SYSTEM Filling2Module (* Module Filling2, generated from its module specification *)
  (* Standard: 61499-2 *)
  APPLICATION Filling2 (* Module Filling2 on target pc (localhost, IO modbus; generated by modgen) *)
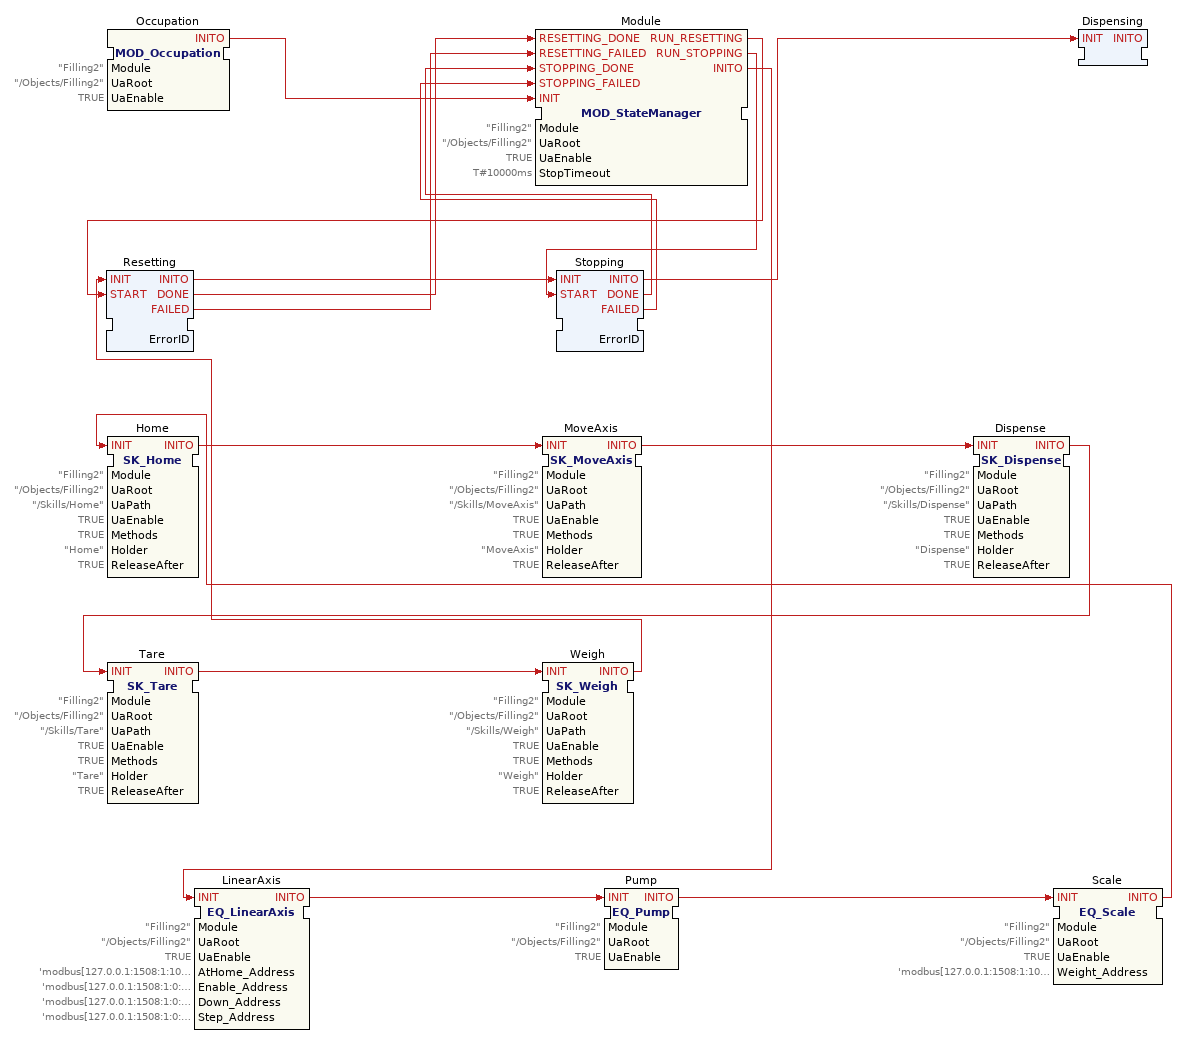
    (* Group ModuleLevel: Module level: occupation, PackML state manager, start-up and the target's IO lines *)
    (* Group ModuleLevelSkills: Module level skills: Control, Sequences (Execute, Stop) of skill primitives and Release; OPC UA /Skills/<name> *)
    (* Group Procedures: Procedures the module state manager runs while Resetting and Stopping *)
    (* Group SkillPrimitives: Skill primitives: one equipment command until a sensor or a time; OPC UA /Skills/<name> *)
    (* Group EquipmentIO: Equipment IO: the only owners of the IO points; skills send them output values over local channels *)
    FBS
      Occupation : modlib::MOD_Occupation(Module := "Filling2", UaRoot := "/Objects/Filling2", UaEnable := TRUE); (* Who may command the module. A client calls Occupy(Session) at /Objects/Filling2/Occupation first; until it calls Release, only commands with that session id are accepted. Every block hears the owner on loc[Filling2/owner]. *) {SET_ATTRIBUTE(GroupName, ModuleLevel)}
      Module : modlib::MOD_StateManager(Module := "Filling2", UaRoot := "/Objects/Filling2", UaEnable := TRUE, StopTimeout := T#10000ms); (* The module's PackML state. The owner calls Reset, Start, Stop, Abort or Clear at /Objects/Filling2/Module; State is at /Objects/Filling2/Module/State and on loc[Filling2/state]. Reset runs the Resetting procedure, Stop the Stopping procedure; skills may be started only in Execute. *) {SET_ATTRIBUTE(GroupName, ModuleLevel)}
      LinearAxis : filling::EQ_LinearAxis(Module := "Filling2", UaRoot := "/Objects/Filling2", UaEnable := TRUE, AtHome_Address := 'modbus[127.0.0.1:1508:1:10:d0:]', Enable_Address := 'modbus[127.0.0.1:1508:1:0::c0]', Down_Address := 'modbus[127.0.0.1:1508:1:0::c1]', Step_Address := 'modbus[127.0.0.1:1508:1:0::h0]'); (* Equipment LinearAxis: Needle lift, a stepper motor through a step and direction driver, with a limit switch at the top (home). The only block that touches its pins (AtHome = modbus[127.0.0.1:1508:1:10:d0:], Enable = modbus[127.0.0.1:1508:1:0::c0], Down = modbus[127.0.0.1:1508:1:0::c1], Step = modbus[127.0.0.1:1508:1:0::h0]). Skills send it what to switch on loc[Filling2/LinearAxis/cmd]; it reports its inputs on loc[Filling2/LinearAxis/state] and at /Objects/Filling2/Equipment/LinearAxis. *) {SET_ATTRIBUTE(GroupName, EquipmentIO)}
      Pump : filling::EQ_Pump(Module := "Filling2", UaRoot := "/Objects/Filling2", UaEnable := TRUE); (* Equipment Pump: Filling pump; none is wired yet, so it has no outputs and dispensing is a time at the station's flow rate. The only block that touches its pins (no pins). Skills send it what to switch on loc[Filling2/Pump/cmd]; it reports its inputs on loc[Filling2/Pump/state] and at /Objects/Filling2/Equipment/Pump. *) {SET_ATTRIBUTE(GroupName, EquipmentIO)}
      Scale : filling::EQ_Scale(Module := "Filling2", UaRoot := "/Objects/Filling2", UaEnable := TRUE, Weight_Address := 'modbus[127.0.0.1:1508:1:10:i0:]'); (* Equipment Scale: Scale; the hardware has none, so the weight is simulated. The only block that touches its pins (Weight = modbus[127.0.0.1:1508:1:10:i0:]). Skills send it what to switch on loc[Filling2/Scale/cmd]; it reports its inputs on loc[Filling2/Scale/state] and at /Objects/Filling2/Equipment/Scale. *) {SET_ATTRIBUTE(GroupName, EquipmentIO)}
      Home : filling::SK_Home(Module := "Filling2", UaRoot := "/Objects/Filling2", UaPath := "/Skills/Home", UaEnable := TRUE, Methods := TRUE, Holder := "Home", ReleaseAfter := TRUE); (* Skill Home, offered on its own: Needle up to the limit switch; from there its position is known, using LinearAxis. A client calls Start (with the parameters), Stop, Abort or Reset at /Objects/Filling2/Skills/Home; State, ErrorID, Parameters and Results are there too. *) {SET_ATTRIBUTE(GroupName, SkillPrimitives)}
      MoveAxis : filling::SK_MoveAxis(Module := "Filling2", UaRoot := "/Objects/Filling2", UaPath := "/Skills/MoveAxis", UaEnable := TRUE, Methods := TRUE, Holder := "MoveAxis", ReleaseAfter := TRUE); (* Skill MoveAxis, offered on its own: Needle to Position, measured down from the limit switch; the direction follows from where it is, using LinearAxis. A client calls Start (with the parameters), Stop, Abort or Reset at /Objects/Filling2/Skills/MoveAxis; State, ErrorID, Parameters and Results are there too. *) {SET_ATTRIBUTE(GroupName, SkillPrimitives)}
      Dispense : filling::SK_Dispense(Module := "Filling2", UaRoot := "/Objects/Filling2", UaPath := "/Skills/Dispense", UaEnable := TRUE, Methods := TRUE, Holder := "Dispense", ReleaseAfter := TRUE); (* Skill Dispense, offered on its own: Dispense a volume at the station's flow rate (open loop, by time, until a pump is wired), using Pump. A client calls Start (with the parameters), Stop, Abort or Reset at /Objects/Filling2/Skills/Dispense; State, ErrorID, Parameters and Results are there too. *) {SET_ATTRIBUTE(GroupName, SkillPrimitives)}
      Tare : filling::SK_Tare(Module := "Filling2", UaRoot := "/Objects/Filling2", UaPath := "/Skills/Tare", UaEnable := TRUE, Methods := TRUE, Holder := "Tare", ReleaseAfter := TRUE); (* Skill Tare, offered on its own: Tare the scale, using Scale. A client calls Start (with the parameters), Stop, Abort or Reset at /Objects/Filling2/Skills/Tare; State, ErrorID, Parameters and Results are there too. *) {SET_ATTRIBUTE(GroupName, SkillPrimitives)}
      Weigh : filling::SK_Weigh(Module := "Filling2", UaRoot := "/Objects/Filling2", UaPath := "/Skills/Weigh", UaEnable := TRUE, Methods := TRUE, Holder := "Weigh", ReleaseAfter := TRUE); (* Skill Weigh, offered on its own: Read the weight, using Scale. A client calls Start (with the parameters), Stop, Abort or Reset at /Objects/Filling2/Skills/Weigh; State, ErrorID, Parameters and Results are there too. *) {SET_ATTRIBUTE(GroupName, SkillPrimitives)}
    END_FBS
    SUBAPPLICATION Resetting (* Procedure the module runs while Resetting *)
      {SET_ATTRIBUTE(GroupName, Procedures)}
      EVENT_INPUT
        INIT : EInit;
        START;
      END_EVENT
      EVENT_OUTPUT
        INITO : EInit;
        DONE;
        FAILED;
      END_EVENT
      VAR_OUTPUT
        ErrorID : UINT;
      END_VAR
      FBS
        Home : filling::SK_Home(Module := "Filling2", UaRoot := "/Objects/Filling2", UaPath := "/Procedures/Resetting/Home", UaEnable := TRUE, Methods := FALSE, Holder := "Procedures/Resetting", ReleaseAfter := TRUE); (* Step 1 of Resetting: runs the skill Home. Its State and ErrorID are at /Objects/Filling2/Procedures/Resetting/Home; it keeps the equipment under the name Procedures/Resetting. *)
        Tare : filling::SK_Tare(Module := "Filling2", UaRoot := "/Objects/Filling2", UaPath := "/Procedures/Resetting/Tare", UaEnable := TRUE, Methods := FALSE, Holder := "Procedures/Resetting", ReleaseAfter := TRUE); (* Step 2 of Resetting: runs the skill Tare. Its State and ErrorID are at /Objects/Filling2/Procedures/Resetting/Tare; it keeps the equipment under the name Procedures/Resetting. *)
        Fail1 : modlib::SKILL_FailMerge; (* Joins the failures of the steps into one (with its error code), so any step's failure ends the sequence. *)
      END_FBS
      EVENT_CONNECTIONS
        Home.SUCCESS TO Tare.START;
        START TO Home.START;
        Tare.SUCCESS TO DONE;
        Home.FAILURE TO Fail1.FAIL_1;
        Tare.FAILURE TO Fail1.FAIL_2;
        Fail1.FAIL TO FAILED;
        INIT TO Home.INIT;
        Tare.INITO TO INITO;
        Home.INITO TO Tare.INIT;
      END_CONNECTIONS
      DATA_CONNECTIONS
        Home.ErrorID TO Fail1.Error1;
        Tare.ErrorID TO Fail1.Error2;
        Fail1.Error TO ErrorID;
      END_CONNECTIONS
    END_SUBAPPLICATION
    SUBAPPLICATION Stopping (* Procedure the module runs while Stopping *)
      {SET_ATTRIBUTE(GroupName, Procedures)}
      EVENT_INPUT
        INIT : EInit;
        START;
      END_EVENT
      EVENT_OUTPUT
        INITO : EInit;
        DONE;
        FAILED;
      END_EVENT
      VAR_OUTPUT
        ErrorID : UINT;
      END_VAR
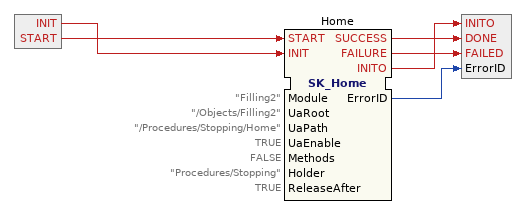
      FBS
        Home : filling::SK_Home(Module := "Filling2", UaRoot := "/Objects/Filling2", UaPath := "/Procedures/Stopping/Home", UaEnable := TRUE, Methods := FALSE, Holder := "Procedures/Stopping", ReleaseAfter := TRUE); (* Step 1 of Stopping: runs the skill Home. Its State and ErrorID are at /Objects/Filling2/Procedures/Stopping/Home; it keeps the equipment under the name Procedures/Stopping. *)
      END_FBS
      EVENT_CONNECTIONS
        START TO Home.START;
        Home.SUCCESS TO DONE;
        Home.FAILURE TO FAILED;
        INIT TO Home.INIT;
        Home.INITO TO INITO;
      END_CONNECTIONS
      DATA_CONNECTIONS
        Home.ErrorID TO ErrorID;
      END_CONNECTIONS
    END_SUBAPPLICATION
    SUBAPPLICATION Dispensing (* Module level skill Dispensing: Needle down, dispense the volume, needle up, weigh (runFillingCycle) *)
      {SET_ATTRIBUTE(GroupName, ModuleLevelSkills)}
      EVENT_INPUT
        INIT : EInit;
      END_EVENT
      EVENT_OUTPUT
        INITO : EInit;
      END_EVENT
      (* Group Core: The skill's state machine: Stop, Abort, Reset, State and ErrorID over OPC UA; gives up everything the skill holds when a run ends *)
      (* Group Start: The Start method: one block per parameter (range check, value for this run), the values published *)
      (* Group Sequences: What the skill does: Execute, and Stop when it is interrupted; private skill primitives in order *)
      (* Group Results: The results published when Execute is done *)
      FBS
        Control : modlib::SKILL_Core(Module := "Filling2", UaRoot := "/Objects/Filling2", UaPath := "/Skills/Dispensing", UaEnable := TRUE, Methods := TRUE, Holder := "Dispensing", ReleaseAll := TRUE); (* The state machine of the skill Dispensing: checks a client's Start (occupation, module in Execute, not running, values in range), publishes State and ErrorID at /Objects/Filling2/Skills/Dispensing, offers Stop, Abort and Reset there, starts Execute and runs Stop when the skill is stopped. *) {SET_ATTRIBUTE(GroupName, Core)}
        UaStart : iec61499::net::SERVER_2_2(QI := TRUE); (* The OPC UA method Start of Dispensing: a client's call (session id and parameters) arrives here; the parameters are checked, then Control answers Accepted or an error code. *) {SET_ATTRIBUTE(GroupName, Start)}
        Volume : modlib::SKILL_Param_LREAL(Default := 1.0, Lower := 0.5, Upper := 10.0); (* The parameter Volume of Dispensing: default 1.0 (Lower 0.5, Upper 10.0); checks a client's value, then holds it for the run and hands it to the steps. *) {SET_ATTRIBUTE(GroupName, Start)}
        PubParams : iec61499::net::PUBLISH_1(QI := TRUE, ID := "opc_ua[WRITE;/Objects/Filling2/Skills/Dispensing/Parameters/Volume]"); (* Writes the parameters of the run to OPC UA: /Objects/Filling2/Skills/Dispensing/Parameters/Volume *) {SET_ATTRIBUTE(GroupName, Start)}
        PubResults : iec61499::net::PUBLISH_1(QI := TRUE, ID := "opc_ua[WRITE;/Objects/Filling2/Skills/Dispensing/Results/Weight]"); (* Writes the results of the run to OPC UA: /Objects/Filling2/Skills/Dispensing/Results/Weight *) {SET_ATTRIBUTE(GroupName, Results)}
      END_FBS
      SUBAPPLICATION Execute (* Dispensing: execute sequence *)
        {SET_ATTRIBUTE(GroupName, Sequences)}
        EVENT_INPUT
          INIT : EInit;
          START;
          HALT;
          ABORT;
          RESET;
        END_EVENT
        EVENT_OUTPUT
          INITO : EInit;
          DONE;
          FAILED;
        END_EVENT
        VAR_INPUT
          Volume : LREAL;
        END_VAR
        VAR_OUTPUT
          ErrorID : UINT;
          Weight : LREAL;
        END_VAR
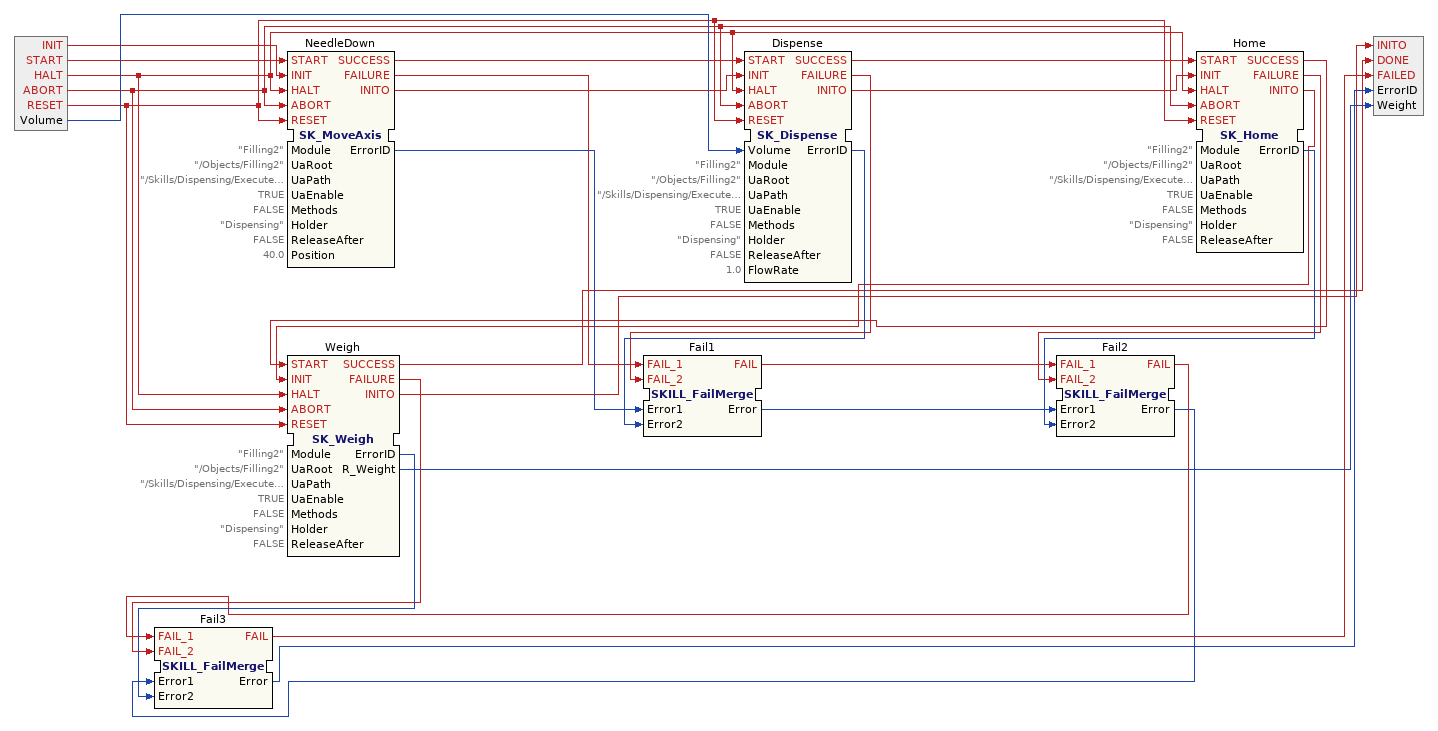
        FBS
          NeedleDown : filling::SK_MoveAxis(Module := "Filling2", UaRoot := "/Objects/Filling2", UaPath := "/Skills/Dispensing/Execute/NeedleDown", UaEnable := TRUE, Methods := FALSE, Holder := "Dispensing", ReleaseAfter := FALSE, Position := 40.0); (* Step 1 of Dispensing / Execute: runs the skill MoveAxis with Position = 40.0. Its State and ErrorID are at /Objects/Filling2/Skills/Dispensing/Execute/NeedleDown; it keeps the equipment under the name Dispensing. *)
          Dispense : filling::SK_Dispense(Module := "Filling2", UaRoot := "/Objects/Filling2", UaPath := "/Skills/Dispensing/Execute/Dispense", UaEnable := TRUE, Methods := FALSE, Holder := "Dispensing", ReleaseAfter := FALSE, FlowRate := 1.0); (* Step 2 of Dispensing / Execute: runs the skill Dispense with FlowRate = 1.0; Volume from Dispensing's Volume. Its State and ErrorID are at /Objects/Filling2/Skills/Dispensing/Execute/Dispense; it keeps the equipment under the name Dispensing. *)
          Home : filling::SK_Home(Module := "Filling2", UaRoot := "/Objects/Filling2", UaPath := "/Skills/Dispensing/Execute/Home", UaEnable := TRUE, Methods := FALSE, Holder := "Dispensing", ReleaseAfter := FALSE); (* Step 3 of Dispensing / Execute: runs the skill Home. Its State and ErrorID are at /Objects/Filling2/Skills/Dispensing/Execute/Home; it keeps the equipment under the name Dispensing. *)
          Weigh : filling::SK_Weigh(Module := "Filling2", UaRoot := "/Objects/Filling2", UaPath := "/Skills/Dispensing/Execute/Weigh", UaEnable := TRUE, Methods := FALSE, Holder := "Dispensing", ReleaseAfter := FALSE); (* Step 4 of Dispensing / Execute: runs the skill Weigh; its Weight is Dispensing's result. Its State and ErrorID are at /Objects/Filling2/Skills/Dispensing/Execute/Weigh; it keeps the equipment under the name Dispensing. *)
          Fail1 : modlib::SKILL_FailMerge; (* Joins the failures of the steps into one (with its error code), so any step's failure ends the sequence. *)
          Fail2 : modlib::SKILL_FailMerge; (* Joins the failures of the steps into one (with its error code), so any step's failure ends the sequence. *)
          Fail3 : modlib::SKILL_FailMerge; (* Joins the failures of the steps into one (with its error code), so any step's failure ends the sequence. *)
        END_FBS
        EVENT_CONNECTIONS
          NeedleDown.SUCCESS TO Dispense.START;
          Dispense.SUCCESS TO Home.START;
          Home.SUCCESS TO Weigh.START;
          START TO NeedleDown.START;
          Weigh.SUCCESS TO DONE;
          NeedleDown.FAILURE TO Fail1.FAIL_1;
          Dispense.FAILURE TO Fail1.FAIL_2;
          Fail1.FAIL TO Fail2.FAIL_1;
          Home.FAILURE TO Fail2.FAIL_2;
          Fail2.FAIL TO Fail3.FAIL_1;
          Weigh.FAILURE TO Fail3.FAIL_2;
          Fail3.FAIL TO FAILED;
          INIT TO NeedleDown.INIT;
          Weigh.INITO TO INITO;
          NeedleDown.INITO TO Dispense.INIT;
          Dispense.INITO TO Home.INIT;
          Home.INITO TO Weigh.INIT;
          HALT TO NeedleDown.HALT;
          HALT TO Dispense.HALT;
          HALT TO Home.HALT;
          HALT TO Weigh.HALT;
          ABORT TO NeedleDown.ABORT;
          ABORT TO Dispense.ABORT;
          ABORT TO Home.ABORT;
          ABORT TO Weigh.ABORT;
          RESET TO NeedleDown.RESET;
          RESET TO Dispense.RESET;
          RESET TO Home.RESET;
          RESET TO Weigh.RESET;
        END_CONNECTIONS
        DATA_CONNECTIONS
          Volume TO Dispense.Volume;
          NeedleDown.ErrorID TO Fail1.Error1;
          Dispense.ErrorID TO Fail1.Error2;
          Fail1.Error TO Fail2.Error1;
          Home.ErrorID TO Fail2.Error2;
          Fail2.Error TO Fail3.Error1;
          Weigh.ErrorID TO Fail3.Error2;
          Fail3.Error TO ErrorID;
          Weigh.R_Weight TO Weight;
        END_CONNECTIONS
      END_SUBAPPLICATION
      SUBAPPLICATION Stop (* Dispensing: stop sequence *)
        {SET_ATTRIBUTE(GroupName, Sequences)}
        EVENT_INPUT
          INIT : EInit;
          START;
          HALT;
          ABORT;
          RESET;
        END_EVENT
        EVENT_OUTPUT
          INITO : EInit;
          DONE;
          FAILED;
        END_EVENT
        VAR_OUTPUT
          ErrorID : UINT;
        END_VAR
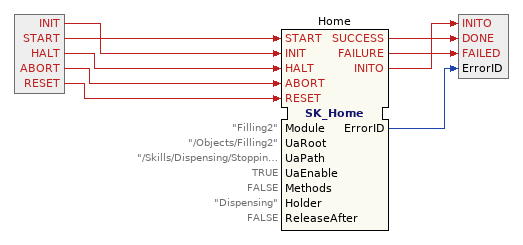
        FBS
          Home : filling::SK_Home(Module := "Filling2", UaRoot := "/Objects/Filling2", UaPath := "/Skills/Dispensing/Stopping/Home", UaEnable := TRUE, Methods := FALSE, Holder := "Dispensing", ReleaseAfter := FALSE); (* Step 1 of Dispensing / Stop: runs the skill Home. Its State and ErrorID are at /Objects/Filling2/Skills/Dispensing/Stopping/Home; it keeps the equipment under the name Dispensing. *)
        END_FBS
        EVENT_CONNECTIONS
          START TO Home.START;
          Home.SUCCESS TO DONE;
          Home.FAILURE TO FAILED;
          INIT TO Home.INIT;
          Home.INITO TO INITO;
          HALT TO Home.HALT;
          ABORT TO Home.ABORT;
          RESET TO Home.RESET;
        END_CONNECTIONS
        DATA_CONNECTIONS
          Home.ErrorID TO ErrorID;
        END_CONNECTIONS
      END_SUBAPPLICATION
      EVENT_CONNECTIONS
        Control.START_RSP TO UaStart.RSP;
        UaStart.IND TO Volume.CHECK;
        Control.RUN TO Volume.LATCH;
        Volume.CHECKED TO Control.START_REQ;
        Volume.LATCHED TO PubParams.REQ;
        PubParams.INITO TO PubParams.REQ;
        Execute.DONE TO PubResults.REQ;
        Volume.LATCHED TO Execute.START;
        Control.HALT_SEQ TO Execute.HALT;
        Control.ABORT_SEQ TO Execute.ABORT;
        Control.RESET_SEQ TO Execute.RESET;
        Execute.DONE TO Control.EXECUTE_DONE;
        Execute.FAILED TO Control.EXECUTE_FAILED;
        Control.RUN_STOPPING TO Stop.START;
        Control.ABORT_SEQ TO Stop.ABORT;
        Control.RESET_SEQ TO Stop.RESET;
        Stop.DONE TO Control.STOPPING_DONE;
        Stop.FAILED TO Control.STOPPING_DONE;
        INIT TO Control.INIT;
        Control.INITO TO UaStart.INIT;
        UaStart.INITO TO Volume.INIT;
        Volume.INITO TO PubParams.INIT;
        PubParams.INITO TO PubResults.INIT;
        PubResults.INITO TO Execute.INIT;
        Execute.INITO TO Stop.INIT;
        Stop.INITO TO INITO;
      END_CONNECTIONS
      DATA_CONNECTIONS
        Control.StartMethodId TO UaStart.ID;
        UaStart.RD_1 TO Control.Session;
        Control.Accepted TO UaStart.SD_1;
        Control.StartError TO UaStart.SD_2;
        UaStart.RD_2 TO Volume.Requested;
        Control.CalledByClient TO Volume.CalledByClient;
        Volume.Value TO PubParams.SD_1;
        Volume.AllInRange TO Control.ParamsInRange;
        Execute.Weight TO PubResults.SD_1;
        Volume.Value TO Execute.Volume;
        Execute.ErrorID TO Control.ExecuteError;
      END_CONNECTIONS
    END_SUBAPPLICATION
    EVENT_CONNECTIONS
      Module.RUN_RESETTING TO Resetting.START;
      Resetting.DONE TO Module.RESETTING_DONE;
      Resetting.FAILED TO Module.RESETTING_FAILED;
      Module.RUN_STOPPING TO Stopping.START;
      Stopping.DONE TO Module.STOPPING_DONE;
      Stopping.FAILED TO Module.STOPPING_FAILED;
      Occupation.INITO TO Module.INIT;
      Module.INITO TO LinearAxis.INIT;
      LinearAxis.INITO TO Pump.INIT;
      Pump.INITO TO Scale.INIT;
      Scale.INITO TO Home.INIT;
      Home.INITO TO MoveAxis.INIT;
      MoveAxis.INITO TO Dispense.INIT;
      Dispense.INITO TO Tare.INIT;
      Tare.INITO TO Weigh.INIT;
      Weigh.INITO TO Resetting.INIT;
      Resetting.INITO TO Stopping.INIT;
      Stopping.INITO TO Dispensing.INIT;
    END_CONNECTIONS
  END_APPLICATION
  APPLICATION Filling2_pi (* Module Filling2 on target pi (192.168.0.173, IO gpio; generated by modgen) *)
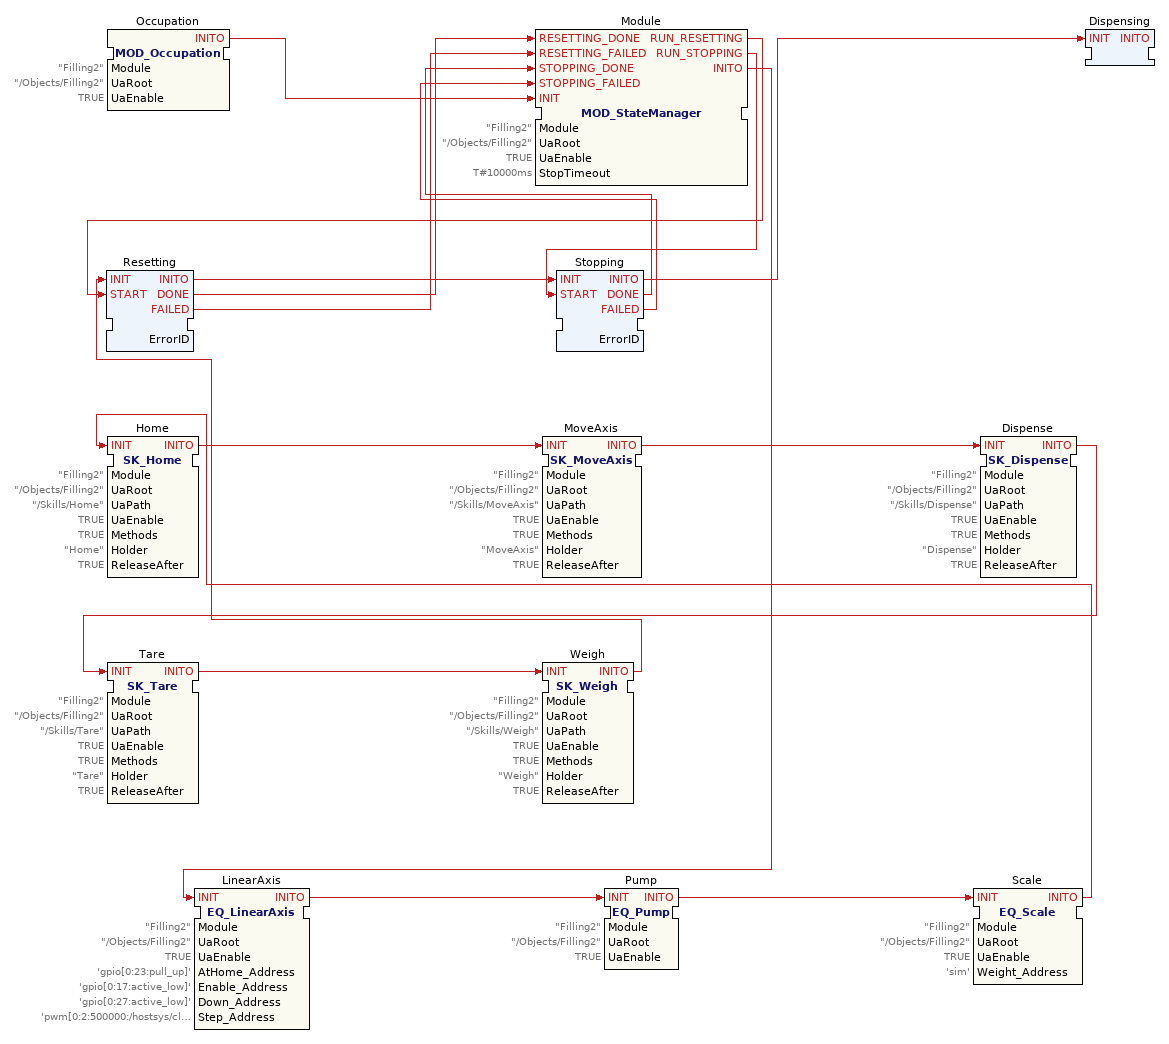
    (* Group ModuleLevel: Module level: occupation, PackML state manager, start-up and the target's IO lines *)
    (* Group ModuleLevelSkills: Module level skills: Control, Sequences (Execute, Stop) of skill primitives and Release; OPC UA /Skills/<name> *)
    (* Group Procedures: Procedures the module state manager runs while Resetting and Stopping *)
    (* Group SkillPrimitives: Skill primitives: one equipment command until a sensor or a time; OPC UA /Skills/<name> *)
    (* Group EquipmentIO: Equipment IO: the only owners of the IO points; skills send them output values over local channels *)
    FBS
      Occupation : modlib::MOD_Occupation(Module := "Filling2", UaRoot := "/Objects/Filling2", UaEnable := TRUE); (* Who may command the module. A client calls Occupy(Session) at /Objects/Filling2/Occupation first; until it calls Release, only commands with that session id are accepted. Every block hears the owner on loc[Filling2/owner]. *) {SET_ATTRIBUTE(GroupName, ModuleLevel)}
      Module : modlib::MOD_StateManager(Module := "Filling2", UaRoot := "/Objects/Filling2", UaEnable := TRUE, StopTimeout := T#10000ms); (* The module's PackML state. The owner calls Reset, Start, Stop, Abort or Clear at /Objects/Filling2/Module; State is at /Objects/Filling2/Module/State and on loc[Filling2/state]. Reset runs the Resetting procedure, Stop the Stopping procedure; skills may be started only in Execute. *) {SET_ATTRIBUTE(GroupName, ModuleLevel)}
      LinearAxis : filling::EQ_LinearAxis(Module := "Filling2", UaRoot := "/Objects/Filling2", UaEnable := TRUE, AtHome_Address := 'gpio[0:23:pull_up]', Enable_Address := 'gpio[0:17:active_low]', Down_Address := 'gpio[0:27:active_low]', Step_Address := 'pwm[0:2:500000:/hostsys/class/pwm]'); (* Equipment LinearAxis: Needle lift, a stepper motor through a step and direction driver, with a limit switch at the top (home). The only block that touches its pins (AtHome = gpio[0:23:pull_up], Enable = gpio[0:17:active_low], Down = gpio[0:27:active_low], Step = pwm[0:2:500000:/hostsys/class/pwm]). Skills send it what to switch on loc[Filling2/LinearAxis/cmd]; it reports its inputs on loc[Filling2/LinearAxis/state] and at /Objects/Filling2/Equipment/LinearAxis. *) {SET_ATTRIBUTE(GroupName, EquipmentIO)}
      Pump : filling::EQ_Pump(Module := "Filling2", UaRoot := "/Objects/Filling2", UaEnable := TRUE); (* Equipment Pump: Filling pump; none is wired yet, so it has no outputs and dispensing is a time at the station's flow rate. The only block that touches its pins (no pins). Skills send it what to switch on loc[Filling2/Pump/cmd]; it reports its inputs on loc[Filling2/Pump/state] and at /Objects/Filling2/Equipment/Pump. *) {SET_ATTRIBUTE(GroupName, EquipmentIO)}
      Scale : filling::EQ_Scale(Module := "Filling2", UaRoot := "/Objects/Filling2", UaEnable := TRUE, Weight_Address := 'sim'); (* Equipment Scale: Scale; the hardware has none, so the weight is simulated. The only block that touches its pins (Weight = sim). Skills send it what to switch on loc[Filling2/Scale/cmd]; it reports its inputs on loc[Filling2/Scale/state] and at /Objects/Filling2/Equipment/Scale. *) {SET_ATTRIBUTE(GroupName, EquipmentIO)}
      Home : filling::SK_Home(Module := "Filling2", UaRoot := "/Objects/Filling2", UaPath := "/Skills/Home", UaEnable := TRUE, Methods := TRUE, Holder := "Home", ReleaseAfter := TRUE); (* Skill Home, offered on its own: Needle up to the limit switch; from there its position is known, using LinearAxis. A client calls Start (with the parameters), Stop, Abort or Reset at /Objects/Filling2/Skills/Home; State, ErrorID, Parameters and Results are there too. *) {SET_ATTRIBUTE(GroupName, SkillPrimitives)}
      MoveAxis : filling::SK_MoveAxis(Module := "Filling2", UaRoot := "/Objects/Filling2", UaPath := "/Skills/MoveAxis", UaEnable := TRUE, Methods := TRUE, Holder := "MoveAxis", ReleaseAfter := TRUE); (* Skill MoveAxis, offered on its own: Needle to Position, measured down from the limit switch; the direction follows from where it is, using LinearAxis. A client calls Start (with the parameters), Stop, Abort or Reset at /Objects/Filling2/Skills/MoveAxis; State, ErrorID, Parameters and Results are there too. *) {SET_ATTRIBUTE(GroupName, SkillPrimitives)}
      Dispense : filling::SK_Dispense(Module := "Filling2", UaRoot := "/Objects/Filling2", UaPath := "/Skills/Dispense", UaEnable := TRUE, Methods := TRUE, Holder := "Dispense", ReleaseAfter := TRUE); (* Skill Dispense, offered on its own: Dispense a volume at the station's flow rate (open loop, by time, until a pump is wired), using Pump. A client calls Start (with the parameters), Stop, Abort or Reset at /Objects/Filling2/Skills/Dispense; State, ErrorID, Parameters and Results are there too. *) {SET_ATTRIBUTE(GroupName, SkillPrimitives)}
      Tare : filling::SK_Tare(Module := "Filling2", UaRoot := "/Objects/Filling2", UaPath := "/Skills/Tare", UaEnable := TRUE, Methods := TRUE, Holder := "Tare", ReleaseAfter := TRUE); (* Skill Tare, offered on its own: Tare the scale, using Scale. A client calls Start (with the parameters), Stop, Abort or Reset at /Objects/Filling2/Skills/Tare; State, ErrorID, Parameters and Results are there too. *) {SET_ATTRIBUTE(GroupName, SkillPrimitives)}
      Weigh : filling::SK_Weigh(Module := "Filling2", UaRoot := "/Objects/Filling2", UaPath := "/Skills/Weigh", UaEnable := TRUE, Methods := TRUE, Holder := "Weigh", ReleaseAfter := TRUE); (* Skill Weigh, offered on its own: Read the weight, using Scale. A client calls Start (with the parameters), Stop, Abort or Reset at /Objects/Filling2/Skills/Weigh; State, ErrorID, Parameters and Results are there too. *) {SET_ATTRIBUTE(GroupName, SkillPrimitives)}
    END_FBS
    SUBAPPLICATION Resetting (* Procedure the module runs while Resetting *)
      {SET_ATTRIBUTE(GroupName, Procedures)}
      EVENT_INPUT
        INIT : EInit;
        START;
      END_EVENT
      EVENT_OUTPUT
        INITO : EInit;
        DONE;
        FAILED;
      END_EVENT
      VAR_OUTPUT
        ErrorID : UINT;
      END_VAR
      FBS
        Home : filling::SK_Home(Module := "Filling2", UaRoot := "/Objects/Filling2", UaPath := "/Procedures/Resetting/Home", UaEnable := TRUE, Methods := FALSE, Holder := "Procedures/Resetting", ReleaseAfter := TRUE); (* Step 1 of Resetting: runs the skill Home. Its State and ErrorID are at /Objects/Filling2/Procedures/Resetting/Home; it keeps the equipment under the name Procedures/Resetting. *)
        Tare : filling::SK_Tare(Module := "Filling2", UaRoot := "/Objects/Filling2", UaPath := "/Procedures/Resetting/Tare", UaEnable := TRUE, Methods := FALSE, Holder := "Procedures/Resetting", ReleaseAfter := TRUE); (* Step 2 of Resetting: runs the skill Tare. Its State and ErrorID are at /Objects/Filling2/Procedures/Resetting/Tare; it keeps the equipment under the name Procedures/Resetting. *)
        Fail1 : modlib::SKILL_FailMerge; (* Joins the failures of the steps into one (with its error code), so any step's failure ends the sequence. *)
      END_FBS
      EVENT_CONNECTIONS
        Home.SUCCESS TO Tare.START;
        START TO Home.START;
        Tare.SUCCESS TO DONE;
        Home.FAILURE TO Fail1.FAIL_1;
        Tare.FAILURE TO Fail1.FAIL_2;
        Fail1.FAIL TO FAILED;
        INIT TO Home.INIT;
        Tare.INITO TO INITO;
        Home.INITO TO Tare.INIT;
      END_CONNECTIONS
      DATA_CONNECTIONS
        Home.ErrorID TO Fail1.Error1;
        Tare.ErrorID TO Fail1.Error2;
        Fail1.Error TO ErrorID;
      END_CONNECTIONS
    END_SUBAPPLICATION
    SUBAPPLICATION Stopping (* Procedure the module runs while Stopping *)
      {SET_ATTRIBUTE(GroupName, Procedures)}
      EVENT_INPUT
        INIT : EInit;
        START;
      END_EVENT
      EVENT_OUTPUT
        INITO : EInit;
        DONE;
        FAILED;
      END_EVENT
      VAR_OUTPUT
        ErrorID : UINT;
      END_VAR
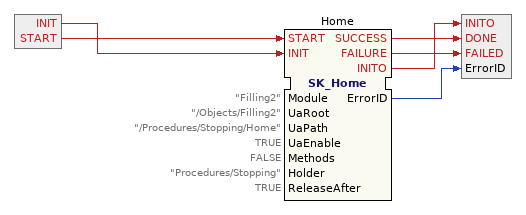
      FBS
        Home : filling::SK_Home(Module := "Filling2", UaRoot := "/Objects/Filling2", UaPath := "/Procedures/Stopping/Home", UaEnable := TRUE, Methods := FALSE, Holder := "Procedures/Stopping", ReleaseAfter := TRUE); (* Step 1 of Stopping: runs the skill Home. Its State and ErrorID are at /Objects/Filling2/Procedures/Stopping/Home; it keeps the equipment under the name Procedures/Stopping. *)
      END_FBS
      EVENT_CONNECTIONS
        START TO Home.START;
        Home.SUCCESS TO DONE;
        Home.FAILURE TO FAILED;
        INIT TO Home.INIT;
        Home.INITO TO INITO;
      END_CONNECTIONS
      DATA_CONNECTIONS
        Home.ErrorID TO ErrorID;
      END_CONNECTIONS
    END_SUBAPPLICATION
    SUBAPPLICATION Dispensing (* Module level skill Dispensing: Needle down, dispense the volume, needle up, weigh (runFillingCycle) *)
      {SET_ATTRIBUTE(GroupName, ModuleLevelSkills)}
      EVENT_INPUT
        INIT : EInit;
      END_EVENT
      EVENT_OUTPUT
        INITO : EInit;
      END_EVENT
      (* Group Core: The skill's state machine: Stop, Abort, Reset, State and ErrorID over OPC UA; gives up everything the skill holds when a run ends *)
      (* Group Start: The Start method: one block per parameter (range check, value for this run), the values published *)
      (* Group Sequences: What the skill does: Execute, and Stop when it is interrupted; private skill primitives in order *)
      (* Group Results: The results published when Execute is done *)
      FBS
        Control : modlib::SKILL_Core(Module := "Filling2", UaRoot := "/Objects/Filling2", UaPath := "/Skills/Dispensing", UaEnable := TRUE, Methods := TRUE, Holder := "Dispensing", ReleaseAll := TRUE); (* The state machine of the skill Dispensing: checks a client's Start (occupation, module in Execute, not running, values in range), publishes State and ErrorID at /Objects/Filling2/Skills/Dispensing, offers Stop, Abort and Reset there, starts Execute and runs Stop when the skill is stopped. *) {SET_ATTRIBUTE(GroupName, Core)}
        UaStart : iec61499::net::SERVER_2_2(QI := TRUE); (* The OPC UA method Start of Dispensing: a client's call (session id and parameters) arrives here; the parameters are checked, then Control answers Accepted or an error code. *) {SET_ATTRIBUTE(GroupName, Start)}
        Volume : modlib::SKILL_Param_LREAL(Default := 1.0, Lower := 0.5, Upper := 10.0); (* The parameter Volume of Dispensing: default 1.0 (Lower 0.5, Upper 10.0); checks a client's value, then holds it for the run and hands it to the steps. *) {SET_ATTRIBUTE(GroupName, Start)}
        PubParams : iec61499::net::PUBLISH_1(QI := TRUE, ID := "opc_ua[WRITE;/Objects/Filling2/Skills/Dispensing/Parameters/Volume]"); (* Writes the parameters of the run to OPC UA: /Objects/Filling2/Skills/Dispensing/Parameters/Volume *) {SET_ATTRIBUTE(GroupName, Start)}
        PubResults : iec61499::net::PUBLISH_1(QI := TRUE, ID := "opc_ua[WRITE;/Objects/Filling2/Skills/Dispensing/Results/Weight]"); (* Writes the results of the run to OPC UA: /Objects/Filling2/Skills/Dispensing/Results/Weight *) {SET_ATTRIBUTE(GroupName, Results)}
      END_FBS
      SUBAPPLICATION Execute (* Dispensing: execute sequence *)
        {SET_ATTRIBUTE(GroupName, Sequences)}
        EVENT_INPUT
          INIT : EInit;
          START;
          HALT;
          ABORT;
          RESET;
        END_EVENT
        EVENT_OUTPUT
          INITO : EInit;
          DONE;
          FAILED;
        END_EVENT
        VAR_INPUT
          Volume : LREAL;
        END_VAR
        VAR_OUTPUT
          ErrorID : UINT;
          Weight : LREAL;
        END_VAR
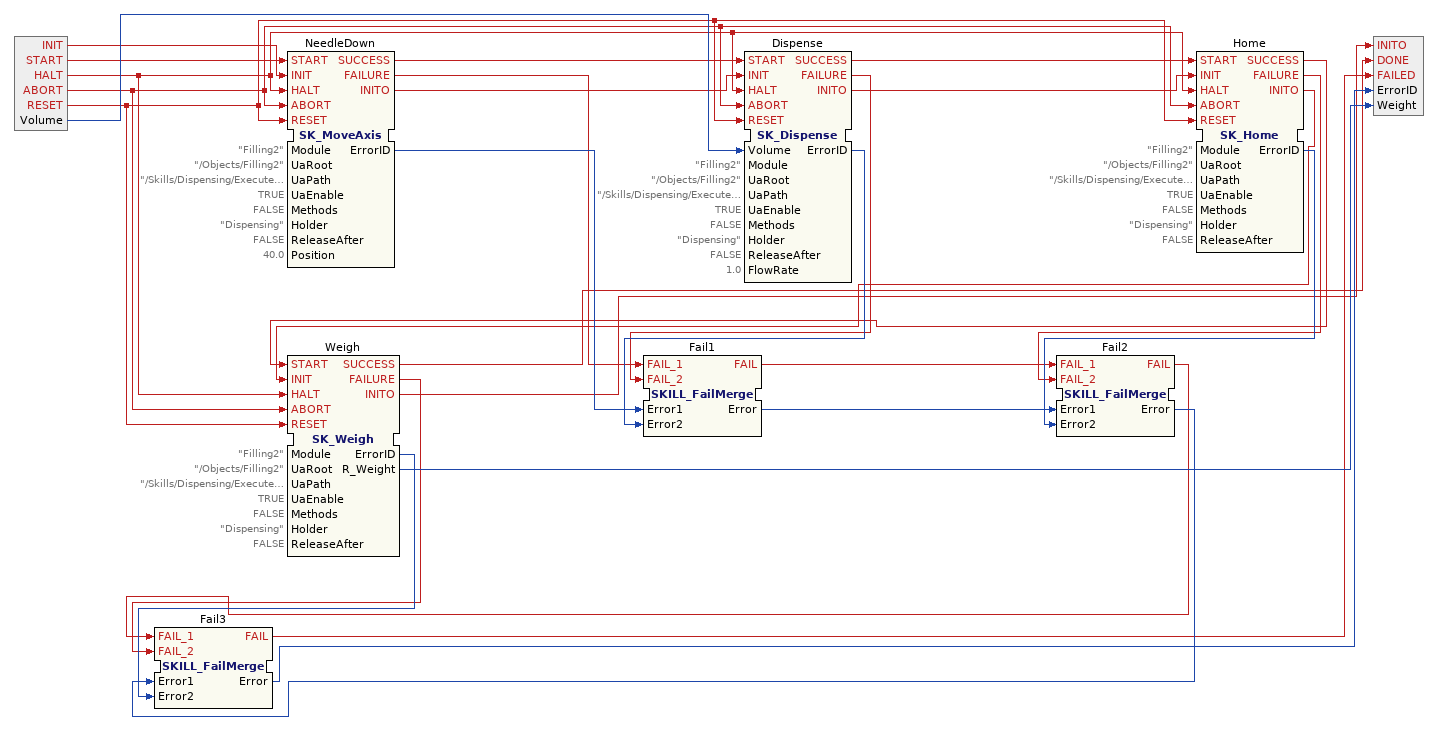
        FBS
          NeedleDown : filling::SK_MoveAxis(Module := "Filling2", UaRoot := "/Objects/Filling2", UaPath := "/Skills/Dispensing/Execute/NeedleDown", UaEnable := TRUE, Methods := FALSE, Holder := "Dispensing", ReleaseAfter := FALSE, Position := 40.0); (* Step 1 of Dispensing / Execute: runs the skill MoveAxis with Position = 40.0. Its State and ErrorID are at /Objects/Filling2/Skills/Dispensing/Execute/NeedleDown; it keeps the equipment under the name Dispensing. *)
          Dispense : filling::SK_Dispense(Module := "Filling2", UaRoot := "/Objects/Filling2", UaPath := "/Skills/Dispensing/Execute/Dispense", UaEnable := TRUE, Methods := FALSE, Holder := "Dispensing", ReleaseAfter := FALSE, FlowRate := 1.0); (* Step 2 of Dispensing / Execute: runs the skill Dispense with FlowRate = 1.0; Volume from Dispensing's Volume. Its State and ErrorID are at /Objects/Filling2/Skills/Dispensing/Execute/Dispense; it keeps the equipment under the name Dispensing. *)
          Home : filling::SK_Home(Module := "Filling2", UaRoot := "/Objects/Filling2", UaPath := "/Skills/Dispensing/Execute/Home", UaEnable := TRUE, Methods := FALSE, Holder := "Dispensing", ReleaseAfter := FALSE); (* Step 3 of Dispensing / Execute: runs the skill Home. Its State and ErrorID are at /Objects/Filling2/Skills/Dispensing/Execute/Home; it keeps the equipment under the name Dispensing. *)
          Weigh : filling::SK_Weigh(Module := "Filling2", UaRoot := "/Objects/Filling2", UaPath := "/Skills/Dispensing/Execute/Weigh", UaEnable := TRUE, Methods := FALSE, Holder := "Dispensing", ReleaseAfter := FALSE); (* Step 4 of Dispensing / Execute: runs the skill Weigh; its Weight is Dispensing's result. Its State and ErrorID are at /Objects/Filling2/Skills/Dispensing/Execute/Weigh; it keeps the equipment under the name Dispensing. *)
          Fail1 : modlib::SKILL_FailMerge; (* Joins the failures of the steps into one (with its error code), so any step's failure ends the sequence. *)
          Fail2 : modlib::SKILL_FailMerge; (* Joins the failures of the steps into one (with its error code), so any step's failure ends the sequence. *)
          Fail3 : modlib::SKILL_FailMerge; (* Joins the failures of the steps into one (with its error code), so any step's failure ends the sequence. *)
        END_FBS
        EVENT_CONNECTIONS
          NeedleDown.SUCCESS TO Dispense.START;
          Dispense.SUCCESS TO Home.START;
          Home.SUCCESS TO Weigh.START;
          START TO NeedleDown.START;
          Weigh.SUCCESS TO DONE;
          NeedleDown.FAILURE TO Fail1.FAIL_1;
          Dispense.FAILURE TO Fail1.FAIL_2;
          Fail1.FAIL TO Fail2.FAIL_1;
          Home.FAILURE TO Fail2.FAIL_2;
          Fail2.FAIL TO Fail3.FAIL_1;
          Weigh.FAILURE TO Fail3.FAIL_2;
          Fail3.FAIL TO FAILED;
          INIT TO NeedleDown.INIT;
          Weigh.INITO TO INITO;
          NeedleDown.INITO TO Dispense.INIT;
          Dispense.INITO TO Home.INIT;
          Home.INITO TO Weigh.INIT;
          HALT TO NeedleDown.HALT;
          HALT TO Dispense.HALT;
          HALT TO Home.HALT;
          HALT TO Weigh.HALT;
          ABORT TO NeedleDown.ABORT;
          ABORT TO Dispense.ABORT;
          ABORT TO Home.ABORT;
          ABORT TO Weigh.ABORT;
          RESET TO NeedleDown.RESET;
          RESET TO Dispense.RESET;
          RESET TO Home.RESET;
          RESET TO Weigh.RESET;
        END_CONNECTIONS
        DATA_CONNECTIONS
          Volume TO Dispense.Volume;
          NeedleDown.ErrorID TO Fail1.Error1;
          Dispense.ErrorID TO Fail1.Error2;
          Fail1.Error TO Fail2.Error1;
          Home.ErrorID TO Fail2.Error2;
          Fail2.Error TO Fail3.Error1;
          Weigh.ErrorID TO Fail3.Error2;
          Fail3.Error TO ErrorID;
          Weigh.R_Weight TO Weight;
        END_CONNECTIONS
      END_SUBAPPLICATION
      SUBAPPLICATION Stop (* Dispensing: stop sequence *)
        {SET_ATTRIBUTE(GroupName, Sequences)}
        EVENT_INPUT
          INIT : EInit;
          START;
          HALT;
          ABORT;
          RESET;
        END_EVENT
        EVENT_OUTPUT
          INITO : EInit;
          DONE;
          FAILED;
        END_EVENT
        VAR_OUTPUT
          ErrorID : UINT;
        END_VAR
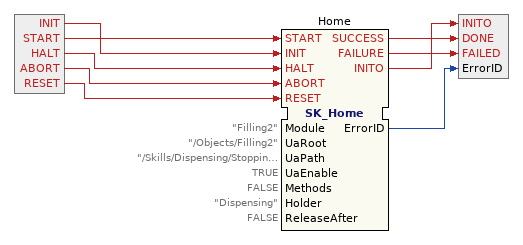
        FBS
          Home : filling::SK_Home(Module := "Filling2", UaRoot := "/Objects/Filling2", UaPath := "/Skills/Dispensing/Stopping/Home", UaEnable := TRUE, Methods := FALSE, Holder := "Dispensing", ReleaseAfter := FALSE); (* Step 1 of Dispensing / Stop: runs the skill Home. Its State and ErrorID are at /Objects/Filling2/Skills/Dispensing/Stopping/Home; it keeps the equipment under the name Dispensing. *)
        END_FBS
        EVENT_CONNECTIONS
          START TO Home.START;
          Home.SUCCESS TO DONE;
          Home.FAILURE TO FAILED;
          INIT TO Home.INIT;
          Home.INITO TO INITO;
          HALT TO Home.HALT;
          ABORT TO Home.ABORT;
          RESET TO Home.RESET;
        END_CONNECTIONS
        DATA_CONNECTIONS
          Home.ErrorID TO ErrorID;
        END_CONNECTIONS
      END_SUBAPPLICATION
      EVENT_CONNECTIONS
        Control.START_RSP TO UaStart.RSP;
        UaStart.IND TO Volume.CHECK;
        Control.RUN TO Volume.LATCH;
        Volume.CHECKED TO Control.START_REQ;
        Volume.LATCHED TO PubParams.REQ;
        PubParams.INITO TO PubParams.REQ;
        Execute.DONE TO PubResults.REQ;
        Volume.LATCHED TO Execute.START;
        Control.HALT_SEQ TO Execute.HALT;
        Control.ABORT_SEQ TO Execute.ABORT;
        Control.RESET_SEQ TO Execute.RESET;
        Execute.DONE TO Control.EXECUTE_DONE;
        Execute.FAILED TO Control.EXECUTE_FAILED;
        Control.RUN_STOPPING TO Stop.START;
        Control.ABORT_SEQ TO Stop.ABORT;
        Control.RESET_SEQ TO Stop.RESET;
        Stop.DONE TO Control.STOPPING_DONE;
        Stop.FAILED TO Control.STOPPING_DONE;
        INIT TO Control.INIT;
        Control.INITO TO UaStart.INIT;
        UaStart.INITO TO Volume.INIT;
        Volume.INITO TO PubParams.INIT;
        PubParams.INITO TO PubResults.INIT;
        PubResults.INITO TO Execute.INIT;
        Execute.INITO TO Stop.INIT;
        Stop.INITO TO INITO;
      END_CONNECTIONS
      DATA_CONNECTIONS
        Control.StartMethodId TO UaStart.ID;
        UaStart.RD_1 TO Control.Session;
        Control.Accepted TO UaStart.SD_1;
        Control.StartError TO UaStart.SD_2;
        UaStart.RD_2 TO Volume.Requested;
        Control.CalledByClient TO Volume.CalledByClient;
        Volume.Value TO PubParams.SD_1;
        Volume.AllInRange TO Control.ParamsInRange;
        Execute.Weight TO PubResults.SD_1;
        Volume.Value TO Execute.Volume;
        Execute.ErrorID TO Control.ExecuteError;
      END_CONNECTIONS
    END_SUBAPPLICATION
    EVENT_CONNECTIONS
      Module.RUN_RESETTING TO Resetting.START;
      Resetting.DONE TO Module.RESETTING_DONE;
      Resetting.FAILED TO Module.RESETTING_FAILED;
      Module.RUN_STOPPING TO Stopping.START;
      Stopping.DONE TO Module.STOPPING_DONE;
      Stopping.FAILED TO Module.STOPPING_FAILED;
      Occupation.INITO TO Module.INIT;
      Module.INITO TO LinearAxis.INIT;
      LinearAxis.INITO TO Pump.INIT;
      Pump.INITO TO Scale.INIT;
      Scale.INITO TO Home.INIT;
      Home.INITO TO MoveAxis.INIT;
      MoveAxis.INITO TO Dispense.INIT;
      Dispense.INITO TO Tare.INIT;
      Tare.INITO TO Weigh.INIT;
      Weigh.INITO TO Resetting.INIT;
      Resetting.INITO TO Stopping.INIT;
      Stopping.INITO TO Dispensing.INIT;
    END_CONNECTIONS
  END_APPLICATION
  DEVICE FORTE_PC : iec61499::system::FORTE_PC(MGR_ID := "localhost:61499" (* Device manager socket ID *))
    {SET_ATTRIBUTE(Profile, HOLOBLOC)}
    RESOURCE RES : iec61499::system::EMB_RES
      EVENT_CONNECTIONS
        START.COLD TO Filling2.Occupation.INIT;
        START.WARM TO Filling2.Occupation.INIT;
      END_CONNECTIONS
    END_RESOURCE
  END_DEVICE
  DEVICE FORTE_PI : iec61499::system::FORTE_PC(MGR_ID := "192.168.0.173:61499" (* Device manager socket ID *))
    {SET_ATTRIBUTE(Profile, HOLOBLOC)}
    RESOURCE RES : iec61499::system::EMB_RES
      EVENT_CONNECTIONS
        START.COLD TO Filling2_pi.Occupation.INIT;
        START.WARM TO Filling2_pi.Occupation.INIT;
      END_CONNECTIONS
    END_RESOURCE
  END_DEVICE
  MAPPINGS
    Filling2.Occupation ON FORTE_PC.RES;
    Filling2.Module ON FORTE_PC.RES;
    Filling2.LinearAxis ON FORTE_PC.RES;
    Filling2.Pump ON FORTE_PC.RES;
    Filling2.Scale ON FORTE_PC.RES;
    Filling2.Home ON FORTE_PC.RES;
    Filling2.MoveAxis ON FORTE_PC.RES;
    Filling2.Dispense ON FORTE_PC.RES;
    Filling2.Tare ON FORTE_PC.RES;
    Filling2.Weigh ON FORTE_PC.RES;
    Filling2.Resetting ON FORTE_PC.RES;
    Filling2.Stopping ON FORTE_PC.RES;
    Filling2.Dispensing ON FORTE_PC.RES;
    Filling2_pi.Occupation ON FORTE_PI.RES;
    Filling2_pi.Module ON FORTE_PI.RES;
    Filling2_pi.LinearAxis ON FORTE_PI.RES;
    Filling2_pi.Pump ON FORTE_PI.RES;
    Filling2_pi.Scale ON FORTE_PI.RES;
    Filling2_pi.Home ON FORTE_PI.RES;
    Filling2_pi.MoveAxis ON FORTE_PI.RES;
    Filling2_pi.Dispense ON FORTE_PI.RES;
    Filling2_pi.Tare ON FORTE_PI.RES;
    Filling2_pi.Weigh ON FORTE_PI.RES;
    Filling2_pi.Resetting ON FORTE_PI.RES;
    Filling2_pi.Stopping ON FORTE_PI.RES;
    Filling2_pi.Dispensing ON FORTE_PI.RES;
  END_MAPPINGS
END_SYSTEM
